// Characterization of FB_MonetTelescopeControl for a stop during a slew, on mock axes (plan step 1, MONETcommonTests README).
// These tests pin what the code does today, with the line of the behaviour in a comment; they are not a specification. Every
// test owns a rig and runs over many PLC cycles (VAR_INST of the method, one Scan() per cycle); TcUnit calls all test methods
// every cycle, so the rigs warm up their clocks in parallel. A step that does not happen within its cycle budget fails the
// test with a message instead of hanging the run. Failed checks are also noted in GVL_Diag.sFailures (printed by Run-Tests.ps1).
FUNCTION_BLOCK MonetStopDuringSlew_Tests EXTENDS TcUnit.FB_TestSuite
VAR
END_VAR

Stop_During_Slew_One_Stop_For_Each_Moving_Axis();
Stop_Drops_The_Moves_In_The_First_Scan_And_Stops_By_The_Second();
Stop_Clears_The_Slew_Keeps_The_Abort_Until_Settled();
Stop_And_Park_Complete_When_An_Axis_Power_Is_Cut_By_An_Interlock();
Stop_During_Slew_Uses_The_Stop_Dynamics();
GoHome_Over_A_Slew_Stops_At_The_Stop_Dynamics();

// #96: one MC_Stop per axis and stop transaction. A slew moves all three axes at once, so all three are stopped, once.
METHOD PRIVATE Stop_During_Slew_One_Stop_For_Each_Moving_Axis
VAR_INST
	rig			: FB_MonetRig;
	nStep		: INT;
	nCycles		: UINT;
	sTest		: STRING(80);
END_VAR
TEST('Stop_During_Slew_One_Stop_For_Each_Moving_Axis');
sTest := 'Stop_During_Slew_One_Stop_For_Each_Moving_Axis: ';
IF nStep >= 90 THEN
	RETURN;
END_IF
rig.Scan();
nCycles := nCycles + 1;
CASE nStep OF
0:	// wait for the clock, then power on
	IF rig.ClockValid THEN
		rig.fbTel.Init();
		nStep := 10;
		nCycles := 0;
	ELSIF nCycles > 2000 THEN
		AssertTrue(Condition := FALSE, Message := 'the astronomical clock never became valid');
		F_Note(bFailed := TRUE, sText := CONCAT(sTest, 'the astronomical clock never became valid'));
		nStep := 99;
		TEST_FINISHED();
	END_IF
10:	// wait until the startup has finished (READY_STATE 1.0), then slew
	IF rig.Online THEN
		rig.fbTel.Slew(fAzimuth := 180.0, fAltitude := 45.0);
		nStep := 20;
		nCycles := 0;
	ELSIF nCycles > 1500 THEN
		AssertTrue(Condition := FALSE, Message := 'the mock telescope did not reach READY_STATE 1.0');
		F_Note(bFailed := TRUE, sText := CONCAT(CONCAT(sTest, 'the mock telescope did not reach READY_STATE 1.0, it is '), LREAL_TO_STRING(rig.fbTel.ReadyState)));
		nStep := 99;
		TEST_FINISHED();
	END_IF
20:	// wait until the slew moves the axes (all three at once)
	IF rig.fbElev.MoveAxis AND rig.fbAzim.MoveAxis AND rig.fbDero.MoveAxis THEN
		AssertTrue(Condition := rig.fbTel.bSlewActive, Message := 'bSlew is set while the slew runs');
		F_Note(bFailed := NOT rig.fbTel.bSlewActive, sText := CONCAT(sTest, 'bSlew is set while the slew runs'));
		nStep := 30;
		nCycles := 0;
	ELSIF nCycles > 300 THEN
		AssertTrue(Condition := FALSE, Message := 'the slew did not start the axis moves');
		F_Note(bFailed := TRUE, sText := CONCAT(sTest, 'the slew did not start the axis moves'));
		nStep := 99;
		TEST_FINISHED();
	END_IF
30:	// let the moves run for a few scans, then stop
	IF nCycles >= 5 THEN
		rig.fbTel.Stop();
		nStep := 40;
		nCycles := 0;
	END_IF
40:	// wait until the stop has settled
	IF NOT rig.fbTel.bStopActive AND rig.fbTel.bStopped AND nCycles > 5 THEN
		AssertEquals_UINT(Expected := 1, Actual := rig.fbElev.nStopEdges, Message := 'elevation: one stop');
		F_Note(bFailed := rig.fbElev.nStopEdges <> 1, sText := CONCAT(sTest, 'elevation: one stop'));
		AssertEquals_UINT(Expected := 1, Actual := rig.fbAzim.nStopEdges, Message := 'azimuth: one stop');
		F_Note(bFailed := rig.fbAzim.nStopEdges <> 1, sText := CONCAT(sTest, 'azimuth: one stop'));
		AssertEquals_UINT(Expected := 1, Actual := rig.fbDero.nStopEdges, Message := 'derotator: one stop');
		F_Note(bFailed := rig.fbDero.nStopEdges <> 1, sText := CONCAT(sTest, 'derotator: one stop'));
		nStep := 99;
		TEST_FINISHED();
	ELSIF nCycles > 400 THEN
		AssertTrue(Condition := FALSE, Message := 'the stop did not settle');
		F_Note(bFailed := TRUE, sText := CONCAT(sTest, 'the stop did not settle'));
		nStep := 99;
		TEST_FINISHED();
	END_IF
END_CASE
END_METHOD

// _StopTelescope (M:1784): one scan does it all: MoveAxis is dropped on all three axes. The stop request itself (StopAxis)
// follows from the stop transaction; pinned here is that it is there by the end of the second scan (still set, the mock
// stop takes 3 scans).
METHOD PRIVATE Stop_Drops_The_Moves_In_The_First_Scan_And_Stops_By_The_Second
VAR_INST
	rig			: FB_MonetRig;
	nStep		: INT;
	nCycles		: UINT;
	sTest		: STRING(80);
END_VAR
TEST('Stop_Drops_The_Moves_In_The_First_Scan_And_Stops_By_The_Second');
sTest := 'Stop_Drops_The_Moves_In_The_First_Scan_And_Stops_By_The_Second: ';
IF nStep >= 90 THEN
	RETURN;
END_IF
rig.Scan();
nCycles := nCycles + 1;
CASE nStep OF
0:	// wait for the clock, then power on
	IF rig.ClockValid THEN
		rig.fbTel.Init();
		nStep := 10;
		nCycles := 0;
	ELSIF nCycles > 2000 THEN
		AssertTrue(Condition := FALSE, Message := 'the astronomical clock never became valid');
		F_Note(bFailed := TRUE, sText := CONCAT(sTest, 'the astronomical clock never became valid'));
		nStep := 99;
		TEST_FINISHED();
	END_IF
10:	// wait until the startup has finished (READY_STATE 1.0), then slew
	IF rig.Online THEN
		rig.fbTel.Slew(fAzimuth := 180.0, fAltitude := 45.0);
		nStep := 20;
		nCycles := 0;
	ELSIF nCycles > 1500 THEN
		AssertTrue(Condition := FALSE, Message := 'the mock telescope did not reach READY_STATE 1.0');
		F_Note(bFailed := TRUE, sText := CONCAT(CONCAT(sTest, 'the mock telescope did not reach READY_STATE 1.0, it is '), LREAL_TO_STRING(rig.fbTel.ReadyState)));
		nStep := 99;
		TEST_FINISHED();
	END_IF
20:	// wait until the slew moves the axes (all three at once)
	IF rig.fbElev.MoveAxis AND rig.fbAzim.MoveAxis AND rig.fbDero.MoveAxis THEN
		AssertTrue(Condition := rig.fbTel.bSlewActive, Message := 'bSlew is set while the slew runs');
		F_Note(bFailed := NOT rig.fbTel.bSlewActive, sText := CONCAT(sTest, 'bSlew is set while the slew runs'));
		nStep := 30;
		nCycles := 0;
	ELSIF nCycles > 300 THEN
		AssertTrue(Condition := FALSE, Message := 'the slew did not start the axis moves');
		F_Note(bFailed := TRUE, sText := CONCAT(sTest, 'the slew did not start the axis moves'));
		nStep := 99;
		TEST_FINISHED();
	END_IF
30:	// let the moves run for a few scans, then stop
	IF nCycles >= 5 THEN
		rig.fbTel.Stop();
		nStep := 40;
		nCycles := 0;
	END_IF
40:	// scan 1 of the stop has just run
	IF nCycles = 1 THEN
		AssertFalse(Condition := rig.fbElev.MoveAxis OR rig.fbAzim.MoveAxis OR rig.fbDero.MoveAxis, Message := 'scan 1 of the stop drops all moves');
		F_Note(bFailed := (rig.fbElev.MoveAxis OR rig.fbAzim.MoveAxis OR rig.fbDero.MoveAxis), sText := CONCAT(sTest, 'scan 1 of the stop drops all moves'));
	ELSIF nCycles = 2 THEN
		AssertTrue(Condition := rig.fbElev.StopAxis AND rig.fbAzim.StopAxis AND rig.fbDero.StopAxis, Message := 'scan 2: all three axes have their stop request');
		F_Note(bFailed := NOT (rig.fbElev.StopAxis AND rig.fbAzim.StopAxis AND rig.fbDero.StopAxis), sText := CONCAT(sTest, 'scan 2: all three axes have their stop request'));
		nStep := 99;
		TEST_FINISHED();
	END_IF
END_CASE
END_METHOD

// Arbitration (M:495-516): a stop during a slew drops bSlew, sets the abort-pending flag (#84) while the axes stop, releases
// both when the stop has settled, and the telescope stays online.
METHOD PRIVATE Stop_Clears_The_Slew_Keeps_The_Abort_Until_Settled
VAR_INST
	rig			: FB_MonetRig;
	nStep		: INT;
	nCycles		: UINT;
	sTest		: STRING(80);
END_VAR
TEST('Stop_Clears_The_Slew_Keeps_The_Abort_Until_Settled');
sTest := 'Stop_Clears_The_Slew_Keeps_The_Abort_Until_Settled: ';
IF nStep >= 90 THEN
	RETURN;
END_IF
rig.Scan();
nCycles := nCycles + 1;
CASE nStep OF
0:	// wait for the clock, then power on
	IF rig.ClockValid THEN
		rig.fbTel.Init();
		nStep := 10;
		nCycles := 0;
	ELSIF nCycles > 2000 THEN
		AssertTrue(Condition := FALSE, Message := 'the astronomical clock never became valid');
		F_Note(bFailed := TRUE, sText := CONCAT(sTest, 'the astronomical clock never became valid'));
		nStep := 99;
		TEST_FINISHED();
	END_IF
10:	// wait until the startup has finished (READY_STATE 1.0), then slew
	IF rig.Online THEN
		rig.fbTel.Slew(fAzimuth := 180.0, fAltitude := 45.0);
		nStep := 20;
		nCycles := 0;
	ELSIF nCycles > 1500 THEN
		AssertTrue(Condition := FALSE, Message := 'the mock telescope did not reach READY_STATE 1.0');
		F_Note(bFailed := TRUE, sText := CONCAT(CONCAT(sTest, 'the mock telescope did not reach READY_STATE 1.0, it is '), LREAL_TO_STRING(rig.fbTel.ReadyState)));
		nStep := 99;
		TEST_FINISHED();
	END_IF
20:	// wait until the slew moves the axes (all three at once)
	IF rig.fbElev.MoveAxis AND rig.fbAzim.MoveAxis AND rig.fbDero.MoveAxis THEN
		AssertTrue(Condition := rig.fbTel.bSlewActive, Message := 'bSlew is set while the slew runs');
		F_Note(bFailed := NOT rig.fbTel.bSlewActive, sText := CONCAT(sTest, 'bSlew is set while the slew runs'));
		nStep := 30;
		nCycles := 0;
	ELSIF nCycles > 300 THEN
		AssertTrue(Condition := FALSE, Message := 'the slew did not start the axis moves');
		F_Note(bFailed := TRUE, sText := CONCAT(sTest, 'the slew did not start the axis moves'));
		nStep := 99;
		TEST_FINISHED();
	END_IF
30:	// let the moves run for a few scans, then stop
	IF nCycles >= 5 THEN
		rig.fbTel.Stop();
		nStep := 40;
		nCycles := 0;
	END_IF
40:
	IF nCycles = 2 THEN
		AssertFalse(Condition := rig.fbTel.bSlewActive, Message := 'the stop dropped bSlew');
		F_Note(bFailed := (rig.fbTel.bSlewActive), sText := CONCAT(sTest, 'the stop dropped bSlew'));
		AssertTrue(Condition := rig.fbTel.bMoveAbortPending, Message := 'bMoveAbortPending is set while the axes stop');
		F_Note(bFailed := NOT (rig.fbTel.bMoveAbortPending), sText := CONCAT(sTest, 'bMoveAbortPending is set while the axes stop'));
	ELSIF NOT rig.fbTel.bStopActive AND rig.fbTel.bStopped AND nCycles > 5 THEN
		AssertFalse(Condition := rig.fbTel.bMoveAbortPending, Message := 'bMoveAbortPending is released with the stop');
		F_Note(bFailed := (rig.fbTel.bMoveAbortPending), sText := CONCAT(sTest, 'bMoveAbortPending is released with the stop'));
		AssertTrue(Condition := rig.fbTel.ReadyState = 1.0, Message := 'the telescope stays online (READY_STATE 1.0)');
		F_Note(bFailed := NOT (rig.fbTel.ReadyState = 1.0), sText := CONCAT(sTest, 'the telescope stays online (READY_STATE 1.0)'));
		nStep := 99;
		TEST_FINISHED();
	ELSIF nCycles > 400 THEN
		AssertTrue(Condition := FALSE, Message := 'the stop did not settle');
		F_Note(bFailed := TRUE, sText := CONCAT(sTest, 'the stop did not settle'));
		nStep := 99;
		TEST_FINISHED();
	END_IF
END_CASE
END_METHOD

// #232 (MONET/S 2026-11-09, MS-158): the brake closes after the elevation was disabled at standstill, and HalfBROT powers the azimuth only
// with the brake open (fbAxis.Enable := bEnable AND bAtRest AND bBrakeOpen), so the NC azimuth goes to Disabled: bEnable (the request)
// stays TRUE, fbAxis.Ready and StandStill are FALSE. bStopped used the request and stayed FALSE for ever: a park and a stop were held
// with no progress and no log line. The mock core models the NC state Disabled with bPowerLost. A stop settles, then a park completes.
METHOD PRIVATE Stop_And_Park_Complete_When_An_Axis_Power_Is_Cut_By_An_Interlock
VAR_INST
	rig			: FB_MonetRig;
	nStep		: INT;
	nCycles		: UINT;
	sTest		: STRING(80);
END_VAR
TEST('Stop_And_Park_Complete_When_An_Axis_Power_Is_Cut_By_An_Interlock');
sTest := 'Stop_And_Park_Complete_When_An_Axis_Power_Is_Cut_By_An_Interlock: ';
IF nStep >= 90 THEN
	RETURN;
END_IF
rig.Scan();
nCycles := nCycles + 1;
CASE nStep OF
0:	// wait for the clock, then power on
	IF rig.ClockValid THEN
		rig.fbTel.Init();
		nStep := 10;
		nCycles := 0;
	ELSIF nCycles > 2000 THEN
		AssertTrue(Condition := FALSE, Message := 'the astronomical clock never became valid');
		F_Note(bFailed := TRUE, sText := CONCAT(sTest, 'the astronomical clock never became valid'));
		nStep := 99;
		TEST_FINISHED();
	END_IF
10:	// online: the azimuth loses its power (request unchanged) and the elevation is disabled, as after the brake interlock
	IF rig.Online THEN
		rig.SetAzimuthPowerLost(TRUE);
		nStep := 20;
		nCycles := 0;
	ELSIF nCycles > 1500 THEN
		AssertTrue(Condition := FALSE, Message := 'the mock telescope did not reach READY_STATE 1.0');
		F_Note(bFailed := TRUE, sText := CONCAT(sTest, 'the mock telescope did not reach READY_STATE 1.0'));
		nStep := 99;
		TEST_FINISHED();
	END_IF
20:	// the precondition of the bug: the request is TRUE, the axis is not powered and not at standstill
	IF nCycles >= 10 THEN
		AssertTrue(Condition := rig.fbAzim.bEnable AND NOT rig.fbAzim.fbAxis.Ready AND NOT rig.fbAzim.fbAxis.StandStill, Message := 'precondition: azimuth requested, not powered, no StandStill');
		F_Note(bFailed := NOT (rig.fbAzim.bEnable AND NOT rig.fbAzim.fbAxis.Ready AND NOT rig.fbAzim.fbAxis.StandStill), sText := CONCAT(sTest, 'precondition: azimuth requested, not powered, no StandStill'));
		AssertTrue(Condition := rig.fbTel.bStopped, Message := 'bStopped is TRUE: an unpowered axis cannot be moving');
		F_Note(bFailed := NOT rig.fbTel.bStopped, sText := CONCAT(sTest, 'bStopped is TRUE: an unpowered axis cannot be moving'));
		rig.fbTel.Stop();
		nStep := 30;
		nCycles := 0;
	END_IF
30:	// the stop settles
	IF NOT rig.fbTel.bStopActive AND rig.fbTel.bStopped AND nCycles > 5 THEN
		AssertTrue(Condition := TRUE, Message := 'the stop settled');
		rig.fbTel.Park();
		nStep := 40;
		nCycles := 0;
	ELSIF nCycles > 300 THEN
		AssertTrue(Condition := FALSE, Message := 'the stop never settled');
		F_Note(bFailed := TRUE, sText := CONCAT(sTest, 'the stop never settled'));
		nStep := 99;
		TEST_FINISHED();
	END_IF
40:	// the park is dispatched and completes
	IF rig.fbTel.bIsParked THEN
		AssertTrue(Condition := rig.fbTel.bIsParked, Message := 'the park completed');
		F_Note(bFailed := NOT rig.fbTel.bIsParked, sText := CONCAT(sTest, 'the park completed'));
		nStep := 99;
		TEST_FINISHED();
	ELSIF nCycles > 1500 THEN
		AssertTrue(Condition := FALSE, Message := 'the park was held (bStopped never TRUE?)');
		F_Note(bFailed := TRUE, sText := CONCAT(sTest, 'the park was held (bStopped never TRUE?)'));
		nStep := 99;
		TEST_FINISHED();
	END_IF
END_CASE
END_METHOD

// #286: the stop command stops every axis at the stop dynamics of stMotion (f*StopDeceleration/f*StopJerk, BROTLib
// SetStopDynamics), not at the NC parameters: with the NC jerk a stop at speed ran on 12-16 deg on MONET/N.
METHOD PRIVATE Stop_During_Slew_Uses_The_Stop_Dynamics
VAR_INST
	rig			: FB_MonetRig;
	nStep		: INT;
	nCycles		: UINT;
	sTest		: STRING(80);
	stCfg		: BROTLib.ST_MotionConfig;
	nEl0		: UINT;
END_VAR
TEST('Stop_During_Slew_Uses_The_Stop_Dynamics');
sTest := 'Stop_During_Slew_Uses_The_Stop_Dynamics: ';
IF nStep >= 90 THEN
	RETURN;
END_IF
IF nStep = 0 AND nCycles = 0 THEN
	stCfg.fAzimuthStopDeceleration := 4.0;
	stCfg.fAzimuthStopJerk := 21.0;
	stCfg.fElevationStopDeceleration := 3.0;
	stCfg.fElevationStopJerk := 22.0;
	stCfg.fDerotatorStopDeceleration := 5.0;
	stCfg.fDerotatorStopJerk := 23.0;
	rig.SetMotion(stValue := stCfg);
END_IF
rig.Scan();
nCycles := nCycles + 1;
CASE nStep OF
0:	// wait for the clock, then power on
	IF rig.ClockValid THEN
		rig.fbTel.Init();
		nStep := 10;
		nCycles := 0;
	ELSIF nCycles > 2000 THEN
		AssertTrue(Condition := FALSE, Message := 'the astronomical clock never became valid');
		F_Note(bFailed := TRUE, sText := CONCAT(sTest, 'the astronomical clock never became valid'));
		nStep := 99;
		TEST_FINISHED();
	END_IF
10:	// online: slew
	IF rig.Online THEN
		rig.fbTel.Slew(fAzimuth := 180.0, fAltitude := 45.0);
		nStep := 20;
		nCycles := 0;
	ELSIF nCycles > 1500 THEN
		AssertTrue(Condition := FALSE, Message := 'the mock telescope did not reach READY_STATE 1.0');
		F_Note(bFailed := TRUE, sText := CONCAT(sTest, 'the mock telescope did not reach READY_STATE 1.0'));
		nStep := 99;
		TEST_FINISHED();
	END_IF
20:	// the slew moves all three axes
	IF rig.fbElev.MoveAxis AND rig.fbAzim.MoveAxis AND rig.fbDero.MoveAxis AND nCycles >= 5 THEN
		nEl0 := rig.fbElev.nStopEdges;
		rig.fbTel.Stop();
		nStep := 30;
		nCycles := 0;
	ELSIF nCycles > 300 THEN
		AssertTrue(Condition := FALSE, Message := 'the slew did not start the axis moves');
		F_Note(bFailed := TRUE, sText := CONCAT(sTest, 'the slew did not start the axis moves'));
		nStep := 99;
		TEST_FINISHED();
	END_IF
30:	// the stop request of the elevation (MC_Stop reads the dynamics at its rising Execute)
	IF rig.fbElev.nStopEdges > nEl0 THEN
		AssertTrue(Condition := rig.fbAzim.fbAxis.StopDeceleration = 4.0 AND rig.fbAzim.fbAxis.StopJerk = 21.0 AND rig.fbElev.fbAxis.StopDeceleration = 3.0 AND rig.fbElev.fbAxis.StopJerk = 22.0 AND rig.fbDero.fbAxis.StopDeceleration = 5.0 AND rig.fbDero.fbAxis.StopJerk = 23.0, Message := 'every axis stops at the stop dynamics of stMotion');
		F_Note(bFailed := NOT (rig.fbAzim.fbAxis.StopDeceleration = 4.0 AND rig.fbAzim.fbAxis.StopJerk = 21.0 AND rig.fbElev.fbAxis.StopDeceleration = 3.0 AND rig.fbElev.fbAxis.StopJerk = 22.0 AND rig.fbDero.fbAxis.StopDeceleration = 5.0 AND rig.fbDero.fbAxis.StopJerk = 23.0), sText := CONCAT(sTest, 'every axis stops at the stop dynamics of stMotion'));
		nStep := 99;
		TEST_FINISHED();
	ELSIF nCycles > 300 THEN
		AssertTrue(Condition := FALSE, Message := 'the elevation was not stopped');
		F_Note(bFailed := TRUE, sText := CONCAT(sTest, 'the elevation was not stopped'));
		nStep := 99;
		TEST_FINISHED();
	END_IF
END_CASE
END_METHOD

// #286: gohome over a running slew stops the axes first (the abort stop, #84), at the stop dynamics of stMotion as well.
METHOD PRIVATE GoHome_Over_A_Slew_Stops_At_The_Stop_Dynamics
VAR_INST
	rig			: FB_MonetRig;
	nStep		: INT;
	nCycles		: UINT;
	sTest		: STRING(80);
	stCfg		: BROTLib.ST_MotionConfig;
	nEl0		: UINT;
END_VAR
TEST('GoHome_Over_A_Slew_Stops_At_The_Stop_Dynamics');
sTest := 'GoHome_Over_A_Slew_Stops_At_The_Stop_Dynamics: ';
IF nStep >= 90 THEN
	RETURN;
END_IF
IF nStep = 0 AND nCycles = 0 THEN
	stCfg.fAzimuthStopDeceleration := 4.0;
	stCfg.fAzimuthStopJerk := 21.0;
	stCfg.fElevationStopDeceleration := 3.0;
	stCfg.fElevationStopJerk := 22.0;
	stCfg.fDerotatorStopDeceleration := 5.0;
	stCfg.fDerotatorStopJerk := 23.0;
	rig.SetMotion(stValue := stCfg);
END_IF
rig.Scan();
nCycles := nCycles + 1;
CASE nStep OF
0:	// wait for the clock, then power on
	IF rig.ClockValid THEN
		rig.fbTel.Init();
		nStep := 10;
		nCycles := 0;
	ELSIF nCycles > 2000 THEN
		AssertTrue(Condition := FALSE, Message := 'the astronomical clock never became valid');
		F_Note(bFailed := TRUE, sText := CONCAT(sTest, 'the astronomical clock never became valid'));
		nStep := 99;
		TEST_FINISHED();
	END_IF
10:	// online: slew
	IF rig.Online THEN
		rig.fbTel.Slew(fAzimuth := 180.0, fAltitude := 45.0);
		nStep := 20;
		nCycles := 0;
	ELSIF nCycles > 1500 THEN
		AssertTrue(Condition := FALSE, Message := 'the mock telescope did not reach READY_STATE 1.0');
		F_Note(bFailed := TRUE, sText := CONCAT(sTest, 'the mock telescope did not reach READY_STATE 1.0'));
		nStep := 99;
		TEST_FINISHED();
	END_IF
20:	// the slew moves all three axes
	IF rig.fbElev.MoveAxis AND rig.fbAzim.MoveAxis AND rig.fbDero.MoveAxis AND nCycles >= 5 THEN
		nEl0 := rig.fbElev.nStopEdges;
		rig.fbTel.Home();
		nStep := 30;
		nCycles := 0;
	ELSIF nCycles > 300 THEN
		AssertTrue(Condition := FALSE, Message := 'the slew did not start the axis moves');
		F_Note(bFailed := TRUE, sText := CONCAT(sTest, 'the slew did not start the axis moves'));
		nStep := 99;
		TEST_FINISHED();
	END_IF
30:	// the stop request of the elevation (MC_Stop reads the dynamics at its rising Execute)
	IF rig.fbElev.nStopEdges > nEl0 THEN
		AssertTrue(Condition := rig.fbAzim.fbAxis.StopDeceleration = 4.0 AND rig.fbAzim.fbAxis.StopJerk = 21.0 AND rig.fbElev.fbAxis.StopDeceleration = 3.0 AND rig.fbElev.fbAxis.StopJerk = 22.0 AND rig.fbDero.fbAxis.StopDeceleration = 5.0 AND rig.fbDero.fbAxis.StopJerk = 23.0, Message := 'every axis stops at the stop dynamics of stMotion');
		F_Note(bFailed := NOT (rig.fbAzim.fbAxis.StopDeceleration = 4.0 AND rig.fbAzim.fbAxis.StopJerk = 21.0 AND rig.fbElev.fbAxis.StopDeceleration = 3.0 AND rig.fbElev.fbAxis.StopJerk = 22.0 AND rig.fbDero.fbAxis.StopDeceleration = 5.0 AND rig.fbDero.fbAxis.StopJerk = 23.0), sText := CONCAT(sTest, 'every axis stops at the stop dynamics of stMotion'));
		nStep := 99;
		TEST_FINISHED();
	ELSIF nCycles > 300 THEN
		AssertTrue(Condition := FALSE, Message := 'the elevation was not stopped');
		F_Note(bFailed := TRUE, sText := CONCAT(sTest, 'the elevation was not stopped'));
		nStep := 99;
		TEST_FINISHED();
	END_IF
END_CASE
END_METHOD

END_FUNCTION_BLOCK

(* stored: Version 1.1.0.1, ProductVersion 3.1.4024.15
   POU MonetStopDuringSlew_Tests: Id {a4fe9a52-989d-4d3e-be2e-00ce5f773a71}, SpecialFunc None
   Method Stop_During_Slew_One_Stop_For_Each_Moving_Axis: Id {16f3a334-4063-405e-93db-2bd09d2218a5}
   Method Stop_Drops_The_Moves_In_The_First_Scan_And_Stops_By_The_Second: Id {8dfec628-3d7a-44af-8920-0ef8fd8d632a}
   Method Stop_Clears_The_Slew_Keeps_The_Abort_Until_Settled: Id {5f87de1a-fd97-421b-8f69-0726be211339}
   Method Stop_And_Park_Complete_When_An_Axis_Power_Is_Cut_By_An_Interlock: Id {2e58537e-0767-4ec2-b7ae-cf0d0ba31918}
   Method Stop_During_Slew_Uses_The_Stop_Dynamics: Id {d63dc9a4-ca0b-4dfc-a91e-6c6648613870}
   Method GoHome_Over_A_Slew_Stops_At_The_Stop_Dynamics: Id {5e342e9a-15c4-4c85-87d3-c1ce68a3eeb7} *)
